DATA_BLOCK "Crane_Control_DB"
{ S7_Optimized_Access := 'TRUE' }
VERSION : 0.1
NON_RETAIN
"Crane_Control"

BEGIN

END_DATA_BLOCK

